(* IEC 61131-3 sources: kns-pump-station/tools/tests/fixtures/sample/src/DUTs/Motor, 3 files *)

(* ---- ST_DeviceSts.dut.st ---- *)
// Общее состояние устройства для HMI/SCADA
TYPE ST_DeviceSts :
STRUCT
    eMode : E_DeviceMode;
    eNamur : E_NamurStatus;
    xFault : BOOL;
END_STRUCT
END_TYPE

(* ---- ST_MotorCmd.dut.st ---- *)
// Команды двигателя от HMI/SCADA
TYPE ST_MotorCmd :
STRUCT
    xStart : BOOL;                                  // пуск
    xStop : BOOL;                                   // стоп
    xAck : BOOL;                                    // квитирование
    eMode : E_DeviceMode := E_DeviceMode.Auto;      // заданный режим
    rSpeedSp_rpm : REAL;                            // уставка скорости
END_STRUCT
END_TYPE

(* ---- ST_MotorSts.dut.st ---- *)
// Состояние двигателя: общее состояние устройства плюс данные привода
TYPE ST_MotorSts EXTENDS ST_DeviceSts :
STRUCT
    xRunning : BOOL;
    rSpeed_rpm : REAL;
    aLastFaults : ARRAY[1..3] OF E_NamurStatus;    // последние отказы
    wsText : WSTRING(80);                           // текст состояния для HMI
END_STRUCT
END_TYPE
